// Répertoire des tables (docs/06 § 2)
{attribute 'pack_mode' := '1'}
TYPE ST_TableDir :
STRUCT
    bUsed : BOOL;
    sName : STRING(40);
    eKind : E_TableKind;
    nStart : INT;               // index de la première instruction dans aInstr
    nLength : INT;
END_STRUCT
END_TYPE

(* stored: Version 1.1.0.1, ProductVersion 3.1.4024.12
   DUT ST_TableDir: Id {ecb4d3dd-d37b-55b9-a706-1df7c58f6a8c} *)
